(* IEC 61131-3 sources: tc3-emulator/examples, 7 files *)

(* ---- functions.st ---- *)
FUNCTION F_Add : DINT
VAR_INPUT
    a, b : DINT;
END_VAR
F_Add := a + b;
END_FUNCTION

FUNCTION F_Increment : DINT
VAR_IN_OUT
    value : DINT;
END_VAR
value := value + 1;
F_Increment := value;
END_FUNCTION

(* ---- real_arrays.st ---- *)
FUNCTION F_Mean : LREAL
VAR_INPUT
    samples : ARRAY[1..4] OF LREAL;
END_VAR
VAR
    i : INT;
END_VAR
FOR i := 1 TO 4 DO
    F_Mean := F_Mean + samples[i];
END_FOR;
F_Mean := F_Mean / 4.0;
END_FUNCTION

FUNCTION F_Scale : BOOL
VAR_INPUT
    factor : REAL;
END_VAR
VAR_IN_OUT
    values : ARRAY[-1..1] OF REAL;
END_VAR
VAR
    i : INT;
END_VAR
FOR i := -1 TO 1 DO
    values[i] := values[i] * factor;
END_FOR;
F_Scale := TRUE;
END_FUNCTION

FUNCTION F_Trace : LREAL
VAR_INPUT
    matrix : ARRAY[-1..0, -1..0] OF LREAL;
END_VAR
F_Trace := matrix[-1, -1] + matrix[0, 0];
END_FUNCTION

(* ---- bits.st ---- *)
FUNCTION_BLOCK FB_DeviceWords
VAR_INPUT
    status : WORD;
    enable : BOOL;
    acknowledge : BOOL;
END_VAR
VAR_IN_OUT
    command : WORD;
END_VAR
VAR_OUTPUT
    ready : BOOL;
    fault : BOOL;
    errorCode : BYTE;
END_VAR
VAR CONSTANT
    cReadyBit : INT := 0;
    cFaultBit : INT := 3;
    cEnableBit : INT := 7;
    cAcknowledgeMask : WORD := WORD#8#100000;
END_VAR
ready := status.cReadyBit;
fault := status.cFaultBit;
errorCode := WORD_TO_BYTE(SHR(status, 8));
command.cEnableBit := enable AND NOT fault;
command := (command AND NOT cAcknowledgeMask)
    OR SEL(acknowledge, WORD#0, cAcknowledgeMask);
END_FUNCTION_BLOCK

FUNCTION F_PackWords : DWORD
VAR_INPUT
    low : WORD;
    high : WORD;
END_VAR
F_PackWords := SHL(WORD_TO_DWORD(high), 16) OR WORD_TO_DWORD(low);
END_FUNCTION

FUNCTION F_HighByte : BYTE
VAR_INPUT
    value : DWORD;
END_VAR
F_HighByte := DWORD_TO_BYTE(SHR(value, 24));
END_FUNCTION

FUNCTION F_RotateMask : BYTE
VAR_INPUT
    mask : BYTE;
END_VAR
F_RotateMask := ROL(mask, 1);
END_FUNCTION

(* ---- standard.st ---- *)
TYPE ST_BatchConfig : STRUCT
    target : WORD := 3;
    releaseDelay : TIME := T#100ms;
    speed : REAL := 10.0;
END_STRUCT END_TYPE

FUNCTION_BLOCK FB_Batch
VAR_INPUT
    sensor : BOOL;
    reset : BOOL;
    config : ST_BatchConfig;
END_VAR
VAR_OUTPUT
    count : WORD;
    targetReached : BOOL;
    release : BOOL;
    speedCommand : INT;
END_VAR
VAR
    edge : R_TRIG;
    counter : CTU;
    reachedLatch : RS;
    releaseTimer : TON;
END_VAR
edge(CLK := sensor);
counter(CU := edge.Q, RESET := reset, PV := config.target, CV => count);
reachedLatch(SET := counter.Q, RESET1 := reset, Q1 => targetReached);
releaseTimer(IN := targetReached, PT := config.releaseDelay, Q => release);
speedCommand := REAL_TO_INT(LIMIT(REAL#0.0, config.speed, REAL#100.0));
END_FUNCTION_BLOCK

FUNCTION F_ConstantTable : DINT
VAR CONSTANT
    cCount : INT := 3;
    cScale : INT := cCount * 2;
END_VAR
VAR
    values : ARRAY[1..cCount] OF INT := [cScale, cScale + 2, cScale + 4];
    index : INT;
END_VAR
FOR index := 1 TO cCount DO
    F_ConstantTable := F_ConstantTable + values[index];
END_FOR;
END_FUNCTION

FUNCTION F_SafeRatio : LREAL
VAR_INPUT
    numerator : LREAL;
    denominator : LREAL;
END_VAR
F_SafeRatio := SEL(denominator <> 0.0, 0.0, numerator / denominator);
END_FUNCTION

(* ---- strings.st ---- *)
(* Latin-1 text handling: no TwinCAT installation or external libraries needed. *)
TYPE ST_TextRecipe : STRUCT
    label : STRING(16);
END_STRUCT END_TYPE

FUNCTION F_AlarmText : STRING(80)
VAR_INPUT
    device : STRING(24);
    code : DINT;
    active : BOOL;
END_VAR
F_AlarmText := CONCAT(device, ': alarm ');
F_AlarmText := CONCAT(F_AlarmText, DINT_TO_STRING(code));
F_AlarmText := CONCAT(F_AlarmText, CONCAT(' [', CONCAT(BOOL_TO_STRING(active), ']')));
END_FUNCTION

FUNCTION F_ParseSpeed : DINT
VAR_INPUT command : STRING(80); END_VAR
VAR_OUTPUT valid : BOOL; END_VAR
VAR CONSTANT prefix : STRING(6) := 'SPEED='; END_VAR
valid := LEFT(command, LEN(prefix)) = prefix AND LEN(command) > LEN(prefix);
IF valid THEN
    (* Malformed or overflowing numbers raise a checked execution error. *)
    F_ParseSpeed := STRING_TO_DINT(MID(command, LEN(command), LEN(prefix) + 1));
END_IF;
END_FUNCTION

FUNCTION_BLOCK FB_SpeedCommand
VAR_INPUT command : STRING(80); END_VAR
VAR_OUTPUT accepted : BOOL; speed : DINT; END_VAR
VAR_TEMP nextSpeed : DINT; END_VAR
nextSpeed := F_ParseSpeed(command := command, valid => accepted);
IF accepted THEN
    speed := nextSpeed;
END_IF;
END_FUNCTION_BLOCK

FUNCTION F_AppendLabel : BOOL
VAR_IN_OUT label : STRING(16); END_VAR
VAR_INPUT suffix : STRING(8); END_VAR
label := CONCAT(label, suffix);
F_AppendLabel := TRUE;
END_FUNCTION

(* ---- timers.st ---- *)
FUNCTION F_AddDelay : TIME
VAR_INPUT
    base : TIME;
END_VAR
F_AddDelay := base + T#250ms;
END_FUNCTION

FUNCTION_BLOCK FB_Timers
VAR_INPUT
    signal : BOOL;
    onDelay : TIME := T#100ms;
    offDelay : TIME := T#200ms;
    pulseWidth : TIME := T#50ms;
END_VAR
VAR_OUTPUT
    delayedOn, delayedOff, pulse : BOOL;
    onElapsed, offElapsed, pulseElapsed : TIME;
END_VAR
VAR
    onTimer : TON;
    offTimer : TOF;
    pulseTimer : TP;
END_VAR
onTimer(IN := signal, PT := onDelay, Q => delayedOn, ET => onElapsed);
offTimer(IN := signal, PT := offDelay, Q => delayedOff, ET => offElapsed);
pulseTimer(IN := signal, PT := pulseWidth, Q => pulse, ET => pulseElapsed);
END_FUNCTION_BLOCK

(* ---- user_types.st ---- *)
TYPE
    E_State : (Idle := 0, Waiting := 10, Running := 20) INT := Idle;
    T_Speed : REAL := 1.5;
    T_Recipe : ARRAY[-1..1] OF ST_Config;
END_TYPE

FUNCTION F_Accelerated : ST_Config
VAR_INPUT
    config : ST_Config;
END_VAR
config.speed := config.speed + 1;
F_Accelerated := config;
END_FUNCTION

FUNCTION F_SetSpeed : BOOL
VAR_IN_OUT
    config : ST_Config;
END_VAR
VAR_INPUT
    speed : T_Speed;
END_VAR
config.speed := speed;
F_SetSpeed := TRUE;
END_FUNCTION

FUNCTION F_Recipe : T_Recipe
VAR
    configs : T_Recipe := [(speed := 2, delay := T#50ms), (speed := 4)];
END_VAR
F_Recipe := configs;
END_FUNCTION

FUNCTION_BLOCK FB_Machine
VAR_INPUT
    start : BOOL;
    config : ST_Config;
END_VAR
VAR_OUTPUT
    state : E_State;
    activeSpeed : REAL;
END_VAR
VAR
    delayTimer : TON;
END_VAR
delayTimer(IN := start AND config.enabled, PT := config.delay);
CASE state OF
    E_State.Idle:
        IF start AND config.enabled THEN state := E_State.Waiting; END_IF;
    E_State.Waiting:
        IF NOT start OR NOT config.enabled THEN
            state := E_State.Idle;
        ELSIF delayTimer.Q THEN
            state := E_State.Running;
        END_IF;
    E_State.Running:
        IF NOT start OR NOT config.enabled THEN state := E_State.Idle; END_IF;
END_CASE;
IF state = E_State.Running THEN
    activeSpeed := config.speed;
ELSE
    activeSpeed := 0;
END_IF;
END_FUNCTION_BLOCK
